// Emplacement d'un mover, publié (docs/06 § 6.3)
{attribute 'pack_mode' := '1'}
TYPE ST_SlotStatus :
STRUCT
    bPresent : BOOL;
    sPartId : STRING(40);
    eStatus : E_PartStatus;
    eVerdict : E_Verdict;
    nOrder : UDINT;
END_STRUCT
END_TYPE

(* stored: Version 1.1.0.1, ProductVersion 3.1.4024.12
   DUT ST_SlotStatus: Id {57a9482a-15ec-5753-802f-8b296490e4e6} *)
